{attribute 'qualified_only'}
{attribute 'to_string'}
TYPE E_Sim_Mode :
(
	eManual	:= 0,	// every signal is set by hand
	eAuto	:= 1,	// one wash cycle
	eQueue	:= 2	// clients of arQueue one after another
);
END_TYPE

(* stored: Version 1.1.0.1, ProductVersion 3.1.4026.20
   DUT E_Sim_Mode: Id {6c1f0a54-2b7e-4f0e-9d3a-1e5b7a90c101} *)
